FUNCTION_BLOCK PartidaComReset (* Partida com reset antes: na subida do comando liga o reset por TempoReset, espera TempoPausa e so entao liga o comando (Sulzer HST: bit 2 Reset, bit 0 Start) *)
  (* Standard: 61499-2 *)
  (* Version 1.3, 10/11/2026, Hidryco, Hidryco, 1.3: cfgResetClique - REQ_RESET (clique de reset na IHM) da o pulso de reset tambem com cfgAtivo = FALSE (Sulzer: reset so no clique, sem reset na partida). 1.2: eventos de saida listados no ECAction (sem isso o runtime nao emite nenhum; o ST so liga/desliga). 1.1: REQ_RESET - na subida do ResetIn (reset do EAE), com o equipamento parado e cfgAtivo, da TempoReset de reset; se houver comando de partida no fim, segue a pausa e a partida. 1.0: sequencia reset -> pausa -> partida (1 s / 1 s). Comando FALSE durante a sequencia aborta (reset e comando em FALSE). cfgAtivo = FALSE: repassa o comando como antes (cada REQ gera CNF_CMD). *)
  PACKAGE SE.Nereda;
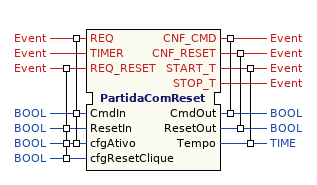
  EVENT_INPUT
    REQ WITH CmdIn, cfgAtivo; (* Novo comando da base (CNF_OUT) *)
    TIMER; (* Fim do tempo (E_DELAY.EO) *)
    REQ_RESET WITH ResetIn, cfgAtivo, cfgResetClique; (* Reset do EAE (ResetCmd) *)
  END_EVENT
  EVENT_OUTPUT
    CNF_CMD WITH CmdOut; (* Comando para a saida (cmdFwd) *)
    CNF_RESET WITH ResetOut; (* Reset para o equipamento *)
    START_T WITH Tempo; (* Inicia o tempo (E_DELAY.START) *)
    STOP_T; (* Cancela o tempo (E_DELAY.STOP) *)
  END_EVENT
  VAR_INPUT
    CmdIn : BOOL; (* Comando da base (OutFwd) *)
    ResetIn : BOOL; (* Reset do EAE (OU de todos os resets do Motor_VS) *)
    cfgAtivo : BOOL; (* TRUE = reset antes de cada partida *)
    cfgResetClique : BOOL; (* TRUE = o clique de reset (REQ_RESET) da o pulso de reset mesmo com cfgAtivo = FALSE *)
  END_VAR
  VAR_OUTPUT
    CmdOut : BOOL; (* Comando para a saida *)
    ResetOut : BOOL; (* Reset para o equipamento *)
    Tempo : TIME; (* Tempo do E_DELAY *)
  END_VAR
  VAR
    fase : INT; (* 0 parado ou repassando, 1 reset, 2 pausa antes da partida, 3 reset pedido pelo EAE *)
    oldResetIn : BOOL; (* ResetIn anterior (borda) *)
    TempoReset : TIME := T#1s; (* Tempo do reset *)
    TempoPausa : TIME := T#1s; (* Pausa entre o fim do reset e a partida *)
  END_VAR
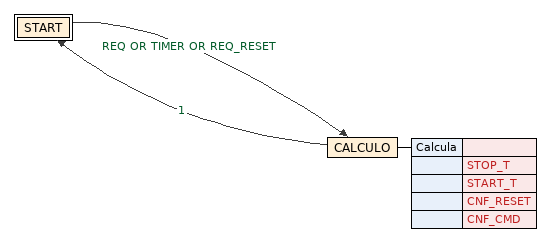
  EC_STATES
    START; (* Estado inicial *)
    CALCULO : Calcula, -> STOP_T, -> START_T, -> CNF_RESET, -> CNF_CMD; (* Calcula; o algoritmo decide quais eventos saem *)
  END_STATES
  EC_TRANSITIONS
    START TO CALCULO := REQ OR TIMER OR REQ_RESET;
    CALCULO TO START := 1;
  END_TRANSITIONS
  ALGORITHM Calcula IN ST: (* Sequencia reset -> pausa -> partida *)
CNF_CMD := FALSE;
CNF_RESET := FALSE;
START_T := FALSE;
STOP_T := FALSE;
IF REQ THEN
    IF NOT CmdIn THEN
        (* parar: aborta a sequencia de partida (o reset pedido pelo EAE, fase 3, termina normalmente) *)
        IF fase = 1 OR fase = 2 THEN
            STOP_T := TRUE;
            fase := 0;
            IF ResetOut THEN
                ResetOut := FALSE;
                CNF_RESET := TRUE;
            END_IF;
        END_IF;
        CmdOut := FALSE;
        CNF_CMD := TRUE;
    ELSIF fase = 0 THEN
        IF cfgAtivo AND NOT CmdOut THEN
            (* partida: primeiro o reset *)
            fase := 1;
            ResetOut := TRUE;
            CNF_RESET := TRUE;
            Tempo := TempoReset;
            START_T := TRUE;
        ELSE
            CmdOut := TRUE;
            CNF_CMD := TRUE;
        END_IF;
    END_IF;
ELSIF REQ_RESET THEN
    (* reset pelo clique: so na subida, parado e sem sequencia em andamento *)
    IF ResetIn AND NOT oldResetIn AND (cfgAtivo OR cfgResetClique) AND fase = 0 AND NOT CmdOut THEN
        fase := 3;
        ResetOut := TRUE;
        CNF_RESET := TRUE;
        Tempo := TempoReset;
        START_T := TRUE;
    END_IF;
    oldResetIn := ResetIn;
ELSIF TIMER THEN
    IF fase = 3 THEN
        ResetOut := FALSE;
        CNF_RESET := TRUE;
        IF CmdIn THEN
            (* chegou comando de partida durante o reset: pausa e parte *)
            fase := 2;
            Tempo := TempoPausa;
            START_T := TRUE;
        ELSE
            fase := 0;
        END_IF;
    ELSIF fase = 1 THEN
        ResetOut := FALSE;
        CNF_RESET := TRUE;
        fase := 2;
        Tempo := TempoPausa;
        START_T := TRUE;
    ELSIF fase = 2 THEN
        fase := 0;
        CmdOut := TRUE;
        CNF_CMD := TRUE;
    END_IF;
END_IF;
  END_ALGORITHM
END_FUNCTION_BLOCK
